(* IEC 61131-3 sources: kns-port-domestic/tools/inventory_tests/fixtures/lib/src/POUs/PsHelper, 1 file *)

(* ---- PsHelper.decl.st ---- *)
// Назначение: имя с префиксом Ps и переменные с именами-ключевыми словами
FUNCTION PsHelper : BOOL
VAR_INPUT
    Override : BOOL;
    Priority : INT;
END_VAR
